Fanuc KAREL source: KA00018.KL

PROGRAM KA00018
%NOLOCKGROUP
VAR
  SRC: REAL
  DST: XYZWPR
BEGIN
  SRC = 2.0
  DST = SRC
END KA00018
